RoboDK station: car_painting 3.rdk

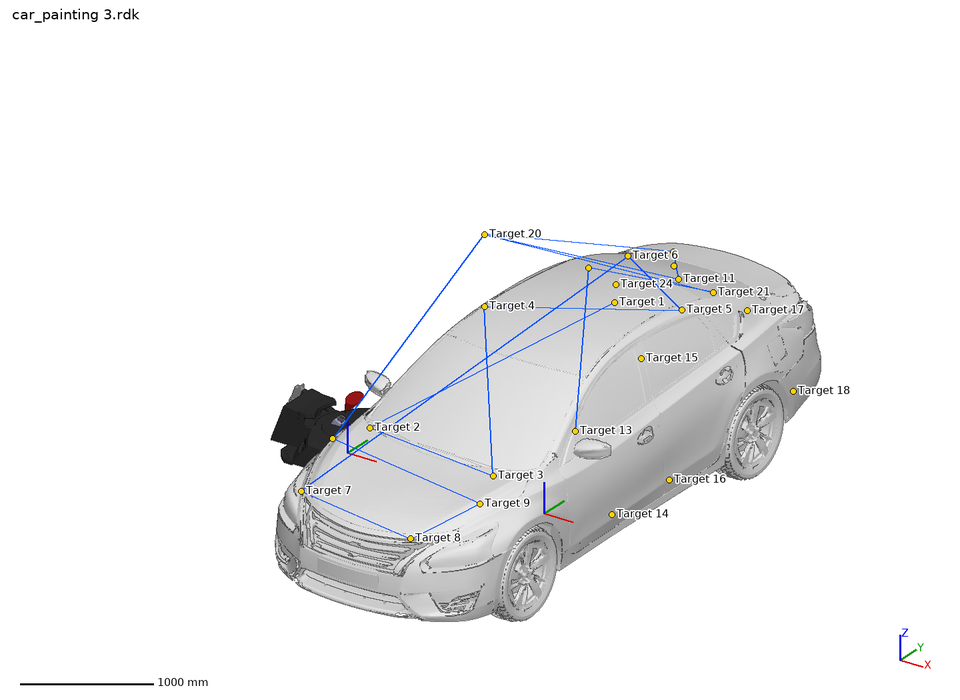
[picture v0: the station drawn from its stored meshes, robots at their saved joint values, targets as dots, program paths as lines]
Station car_painting 3 (saved by RoboDK 6.0.7). Poses are relative to the parent item; angles as X-Y-Z fixed-axis rotations.
  - frame KUKA KR 210 R3100 ultra Base at (0, 0, 0) mm
    - robot KUKA KR 210 R3100 ultra: 6 axes
        joint limits [-185, -140, -120, -350, -122.5, -350] to [185, -5, 155, 350, 122.5, 350]; home [0, -90, 90, 0, 0, 0]; saved at [-29.424, -52.78, 24.902, 2.57, 94.197, 1.598]
      - tool Generic Paint Sprayer, TCP at (50, 0, 700) mm, rotated rx 0 ry 30 rz 0 deg, size 277.6 x 203.2 x 501.7 mm
      - tool Paint Nozzle, TCP at (0, 0, 200) mm, rotated rx 180 ry 0 rz 0 deg
  - program Prog1 (19 instructions, listed below)
  - frame Car_Frame at (1800, 0, 0) mm
    - object Nissan Altima 2013 at (0, 0, 0) mm, size 2245.8 x 5200.8 x 1590 mm, geometry from Nissan Altima 2013.stl
    - target Target 1 (Cartesian target) at (640, 0, 1934) mm, rotated rx -180 ry 0 rz -180 deg; joints [0, -66.141, 36.954, 0, 89.187, 0] of KUKA KR 210 R3100 ultra
    - target Target 2 (Cartesian target) at (-638.65, -1364.5, 1079.42) mm, rotated rx 174.56 ry 3.25 rz -170.84 deg; joints [60.399, -90.418, 102.953, -34.541, 72.996, 77.319] of KUKA KR 210 R3100 ultra
    - target Target 3 (Cartesian target) at (569.96, -1483.73, 1064.93) mm, rotated rx 171.48 ry 0.88 rz -170.48 deg; joints [38.04, -48.846, 47.805, -28.606, 76.343, 48.568] of KUKA KR 210 R3100 ultra
    - target Target 4 (Cartesian target) at (-582.04, 47.56, 1544.2) mm, rotated rx -150.72 ry 0.03 rz -139.53 deg; joints [-6.003, -131.612, 113.224, 4.089, 67.618, 42.32] of KUKA KR 210 R3100 ultra
    - target Target 5 (Cartesian target) at (485.68, 1100.97, 1390.68) mm, rotated rx -166.55 ry -14.54 rz -154.98 deg; joints [-30.565, -60.833, 41.108, 13.15, 94.618, 2.427] of KUKA KR 210 R3100 ultra
    - target Target 6 (Cartesian target) at (-451.98, 1738.11, 1324.58) mm, rotated rx -157.72 ry -3.42 rz -150.29 deg; joints [-64.767, -78.284, 71.355, 31.983, 85.443, -27.718] of KUKA KR 210 R3100 ultra
    - target Target 7 (Cartesian target) at (-755.4, -2100.48, 812.75) mm, rotated rx -157.72 ry -3.42 rz -150.29 deg; joints [74.523, -73.496, 86.549, 145.765, -67.088, -58.208] of KUKA KR 210 R3100 ultra
    - target Target 8 (Cartesian target) at (435.21, -2365.39, 853.53) mm, rotated rx -157.72 ry -3.42 rz -150.29 deg; joints [50.551, -23.508, 12.25, 156.42, -76.689, -92.645] of KUKA KR 210 R3100 ultra
    - target Target 9 (Cartesian target) at (695.7, -1837.37, 1007.74) mm, rotated rx -157.72 ry -3.42 rz -150.29 deg; joints [39.417, -40.307, 36.481, 160.47, -65.722, -100.609] of KUKA KR 210 R3100 ultra
    - target Target 10 (Cartesian target) at (-865.06, -1527.11, 990.04) mm, rotated rx -157.72 ry -3.42 rz -150.29 deg; joints [68.046, -94.782, 111.294, 145.695, -60.704, -61.804] of KUKA KR 210 R3100 ultra
    - target Target 11 (Cartesian target) at (178.8, 1500.41, 1403.06) mm, rotated rx -174.15 ry -4.43 rz -150.4 deg; joints [-40.715, -71.63, 57.081, 189.925, -80.308, -188.903] of KUKA KR 210 R3100 ultra
    - target Target 12 (Cartesian target) at (-359.52, 2197.25, 1202.11) mm, rotated rx -170.21 ry -1.52 rz -149.89 deg; joints [-64.307, -63.206, 54.973, 203.382, -79.356, -211.955] of KUKA KR 210 R3100 ultra
    - target Target 13 (Cartesian target) at (792.65, -730, 1194.78) mm, rotated rx -157.72 ry 0.42 rz -150.29 deg; joints [17.97, -72.117, 70.1, -10.594, 56.299, 56.688] of KUKA KR 210 R3100 ultra
    - target Target 14 (Cartesian target) at (1250.11, -906.27, 700.96) mm, rotated rx -157.72 ry 0.42 rz -150.29 deg; joints [18.543, -47.197, 53.366, -12.261, 48.387, 59.444] of KUKA KR 210 R3100 ultra
    - target Target 15 (Cartesian target) at (709.14, 254.02, 1385.86) mm, rotated rx -157.72 ry 0.42 rz -150.29 deg; joints [-8.226, -72.853, 71.39, 8.418, 55.225, 24.903] of KUKA KR 210 R3100 ultra
    - target Target 16 (Cartesian target) at (960.42, 258.34, 445.14) mm, rotated rx -157.72 ry 0.42 rz -150.29 deg; joints [-7.469, -51.43, 80.281, 15.235, 25.332, 16.51] of KUKA KR 210 R3100 ultra
    - target Target 17 (Cartesian target) at (733.12, 1599.78, 1256.09) mm, rotated rx -157.72 ry 0.42 rz -150.29 deg; joints [-37.551, -43.43, 32.43, 24.375, 72.801, -3.259] of KUKA KR 210 R3100 ultra
    - target Target 18 (Cartesian target) at (961.43, 1880.74, 535.82) mm, rotated rx -157.72 ry 60.42 rz -150.29 deg; joints [-40.295, -27.886, 58.516, -46.206, -43.415, 49.228] of KUKA KR 210 R3100 ultra
    - target Target 20 (Cartesian target) at (-582.04, 47.56, 2144.2) mm, rotated rx -150.72 ry 0.03 rz -139.53 deg; joints [-7.497, -119.703, 70.792, 4.805, 98.145, 43.427] of KUKA KR 210 R3100 ultra
    - target Target 21 (Cartesian target) at (620.53, 1315.55, 1488.37) mm, rotated rx -177.07 ry -6.35 rz -150.64 deg; joints [-29.424, -52.78, 24.902, 2.57, 94.197, 1.598] of KUKA KR 210 R3100 ultra
    - target Target 22 (Cartesian target) at (-335.05, 1052.3, 1532.87) mm, rotated rx -171.84 ry 1 rz -149.58 deg; joints [-42.289, -103.568, 86.635, 13.378, 77.832, -9.168] of KUKA KR 210 R3100 ultra
    - target Target 23 (Cartesian target) at (0.11, 1692.85, 1386.55) mm, rotated rx -163.63 ry -4.97 rz -151.33 deg; joints [-51.523, -68.72, 54.985, 23.065, 85.263, -15.926] of KUKA KR 210 R3100 ultra
    - target Target 24 (Cartesian target) at (39.24, 881.03, 1567.9) mm, rotated rx -174.34 ry -1.31 rz -150.97 deg; joints [-27.642, -92.835, 75.029, 4.309, 78.929, 3.231] of KUKA KR 210 R3100 ultra
  - Python program SprayOn (listed below)
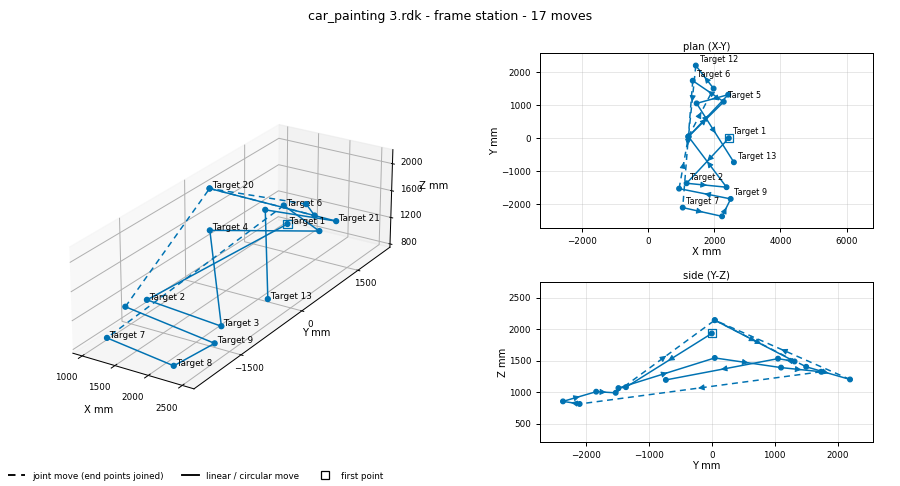
[picture p0: tool path of car_painting 3.rdk in frame station, 17 of 17 moves have a stored position in this frame; points joined in program order, loops and branches not executed]

--- program Prog1 (robot KUKA KR 210 R3100 ultra) ---
  MoveJ (Target 1)
  Call SprayOn(1)
  Set speed (100.0 mm/s)
  MoveL (Target 2)
  MoveL (Target 3)
  MoveL (Target 4)
  MoveL (Target 5)
  MoveL (Target 6)
  MoveJ (Target 7)
  MoveL (Target 8)
  MoveL (Target 9)
  MoveL (Target 10)
  MoveJ (Target 20)
  MoveJ (Target 11)
  MoveL (Target 12)
  MoveJ (Target 20)
  MoveL (Target 21)
  MoveL (Target 22)
  MoveL (Target 13)

--- Python program SprayOn ---
from robodk.robolink import *
from robodk.robomath import *
RDK = Robolink()

tool = RDK.Item('Generic Paint Sprayer', ITEM_TYPE_TOOL)
obj = RDK.Item('Nissan Altima 2013', ITEM_TYPE_OBJECT)

RDK.Spray_Clear()

# Using 50mm cubes limits the "itching" slightly while still overlapping
options = "PROJECT PARTICLE=CUBE(50,50,50) STEP=6x6"

# The 800s make the spray cone massive enough to hit every curve
close_p = [0, 0, 0,    100, 0, 0,    0, 100, 0,    0, 1, 0, 1]
far_p   = [0, 0, 1000, 800, 0, 0,    0, 800, 0,    0, 1, 0, 1]

RDK.Spray_Add(tool, obj, options, Mat([close_p, far_p]).tr())
RDK.Spray_SetState(SPRAY_ON)
